(* IEC 61131-3 sources: guidance-for-physical-ai-production-designer-on-aws/source/plan2cell/crates/plan2cell/tests/fixtures/deploy_check/scene_fit/plc/codesys/head/GVL, 1 file *)

(* ---- GVL_Cell.st ---- *)
(*
 * GVL_Cell - generated by bt2plc 0.1.0 - DO NOT EDIT
 * Plan   : bt_1792156523_scene_fit (cell scene_fit)
 * Grants : planned ticket order
 * IL01   : R1#1 W02 > R2#2 W03 > R1#3 HOME
 * IL02   : R2#1 W01 > R1#2 W04 > R2#3 HOME
 *)
{attribute 'qualified_only'}
VAR_GLOBAL CONSTANT
    (* ========================================================================
       DIMENSIONS (array bounds are literals; *_DIM >= 1)
       ======================================================================== *)
    N_ROBOTS                : INT := 2;
    N_ZONES                 : INT := 2;
    N_OPS                   : INT := 6;
    N_PREDS                 : INT := 0;

    (* ========================================================================
       PROTOCOL / TIMING
       ======================================================================== *)
    PLAN_ID                 : WORD := WORD#16#A1BE;             (* fold of the plan fingerprint *)
    PROD_FOLGE              : WORD := WORD#11;                  (* default production Folge *)
    HOME_FOLGE              : WORD := WORD#125;                 (* blind homing *)
    JOB_NUMBER_BYTE         : BOOL := TRUE;                     (* FALSE: WORD LE bytes 2-3, TRUE: byte 2 *)
    PROFILE_VW              : BOOL := TRUE;                     (* TRUE: VW KS24 signal map and Folge handshake instead of the simulator telegram *)
    GRANT_POLICY            : E_GrantPolicy := E_GrantPolicy.GP_PLANNED;
    HOME_SEQUENTIAL         : BOOL := TRUE;
    AUTO_RUN                : BOOL := TRUE;                     (* start the next cycle automatically *)
    STEP_BYTE               : INT := 4;                         (* robot -> PLC, WORD LE op index *)
    REQ_BYTE                : INT := 28;                        (* robot -> PLC, DWORD LE zone requests *)
    GRANT_BYTE              : INT := 12;                        (* PLC -> robot, DWORD LE zone grants *)
    PLAN_ID_BYTE            : INT := 0;                         (* PLC -> robot, WORD LE plan id *)
    PERMIT_MASK             : DWORD := DWORD#16#80000000;       (* bit 31: permit predecessors *)
    T_RESET_PULSE           : TIME := T#1S;
    T_START_PULSE           : TIME := T#500MS;
    T_STOP_PULSE            : TIME := T#1S;
    T_HANDSHAKE             : TIME := T#5S;
    T_BRINGUP_LIMIT         : TIME := T#1M;                     (* safety enable: PROFINET connection set-up *)
    T_MISMATCH_DEBOUNCE     : TIME := T#200MS;
    T_STOP_DEBOUNCE         : TIME := T#200MS;                  (* job running: ProgRunning and ProgFinished low this long = robot stopped *)
    T_CYCLE_PAUSE           : TIME := T#2S;
    T_START_LIMIT           : TIME := T#15S;
    T_ABORT_LIMIT           : TIME := T#10S;
    T_HOME_LIMIT            : TIME := T#15S500MS;

    (* ========================================================================
       VW KS24 SIGNAL INDICES (used when PROFILE_VW; $IN/$OUT index, 1-based)
       ======================================================================== *)
    VW_READY_OUT            : INT := 9;                         (* O_R_Bereit *)
    VW_RK100_OUT            : INT := 10;                        (* O_R_RK100 safety circuit *)
    VW_AUTO_OUT             : INT := 12;                        (* O_R_Auto *)
    VW_ESTOP_OUT            : INT := 13;                        (* O_R_Notaus *)
    VW_END_OUT              : INT := 14;                        (* O_R_F_ENDE / LPKT *)
    VW_PF0_OUT              : INT := 15;                        (* O_R_PFO home position *)
    VW_STEP_OUT             : INT := 97;                        (* P_PktNr_SPS op index (16 bits) *)
    VW_REL_OUT              : INT := 41;                        (* interlock releases A41-56 *)
    VW_REQ_OUT              : INT := 81;                        (* interlock requests A81-96 *)
    VW_ERR_OUT              : INT := 225;                       (* VW_FEH_BIN_A error code (8 bits) *)
    VW_DRIVES_IN            : INT := 10;                        (* I_R_Ant_Ein *)
    VW_SRB_IN               : INT := 9;                         (* I_R_SRB Folge start *)
    VW_RESET_IN             : INT := 26;                        (* I_R_Quit_St acknowledge *)
    anInterlock             : ARRAY[1..4] OF INT := [1,2,1,2];  (* robot r, zone z -> VW interlock 1..16 (0 = not a member): index (r-1)*2+z *)

    (* ========================================================================
       ROBOTS (index = BT order)
       ======================================================================== *)
    asRobotTag              : ARRAY[1..2] OF STRING(16) := ['R1', 'R2'];
    asRobotNs               : ARRAY[1..2] OF STRING(32) := ['robot1', 'robot2'];
    abRobotActive           : ARRAY[1..2] OF BOOL := [TRUE, TRUE];
    abSafetyBypass          : ARRAY[1..2] OF BOOL := [FALSE, FALSE];(* SIMULATION ONLY: PROFIsafe slot-1 bits not required ([[robot]] safety_bypass) *)
    awRobotProdFolge        : ARRAY[1..2] OF WORD := [WORD#11, WORD#11];
    anRobotFirstOp          : ARRAY[1..2] OF INT := [1, 4];     (* op k of robot r: aOps[anRobotFirstOp[r] + k - 1] *)
    anRobotOpCount          : ARRAY[1..2] OF INT := [3, 3];

    (* ========================================================================
       ZONES - tickets of zone z: aTickets[anZoneFirst[z] .. anZoneFirst[z] + anZoneCount[z] - 1]
       ======================================================================== *)
    asZoneName              : ARRAY[1..2] OF STRING(8) := ['IL01', 'IL02'];
    anZoneFirst             : ARRAY[1..2] OF INT := [1, 4];
    anZoneCount             : ARRAY[1..2] OF INT := [3, 3];
    aTickets                : ARRAY[1..6] OF ST_Ticket := [
        (nRobot := 1, nOp := 1),    (* IL01 R1 #1 W02 *)
        (nRobot := 2, nOp := 2),    (* R2 #2 W03 *)
        (nRobot := 1, nOp := 3),    (* R1 #3 HOME *)
        (nRobot := 2, nOp := 1),    (* IL02 R2 #1 W01 *)
        (nRobot := 1, nOp := 2),    (* R1 #2 W04 *)
        (nRobot := 2, nOp := 3)    (* R2 #3 HOME *)
    ];

    (* ========================================================================
       OPS - op k of robot r: aOps[anRobotFirstOp[r] + k - 1]
       ======================================================================== *)
    (* tLimit = 1.5 x tExpected + 5 s ; tZoneDeadline = 1.5 x ASAP grant + (5 + 0.2) s x depth + 10 s *)
    aOps                    : ARRAY[1..6] OF ST_OpInfo := [
        (nRobot := 1, nOp := 1, dwZoneMask := DWORD#16#00000001, nPredFirst := 0, nPredCount := 0, tExpected := T#7S408MS, tLimit := T#16S112MS, tZoneDeadline := T#10S, sName := 'W02'),    (* R1 #1 W02 *)
        (nRobot := 1, nOp := 2, dwZoneMask := DWORD#16#00000002, nPredFirst := 0, nPredCount := 0, tExpected := T#5S118MS, tLimit := T#12S677MS, tZoneDeadline := T#33S680MS, sName := 'W04'),    (* R1 #2 W04 *)
        (nRobot := 1, nOp := 3, dwZoneMask := DWORD#16#00000001, nPredFirst := 0, nPredCount := 0, tExpected := T#4S522MS, tLimit := T#11S783MS, tZoneDeadline := T#46S557MS, sName := 'HOME'),    (* R1 #3 HOME *)
        (nRobot := 2, nOp := 1, dwZoneMask := DWORD#16#00000002, nPredFirst := 0, nPredCount := 0, tExpected := T#12S320MS, tLimit := T#23S480MS, tZoneDeadline := T#10S, sName := 'W01'),    (* R2 #1 W01 *)
        (nRobot := 2, nOp := 2, dwZoneMask := DWORD#16#00000001, nPredFirst := 0, nPredCount := 0, tExpected := T#5S117MS, tLimit := T#12S676MS, tZoneDeadline := T#33S680MS, sName := 'W03'),    (* R2 #2 W03 *)
        (nRobot := 2, nOp := 3, dwZoneMask := DWORD#16#00000002, nPredFirst := 0, nPredCount := 0, tExpected := T#10S293MS, tLimit := T#20S440MS, tZoneDeadline := T#46S557MS, sName := 'HOME')    (* R2 #3 HOME *)
    ];

    (* ========================================================================
       PERMIT PREDECESSORS - op preds: aPreds[nPredFirst .. nPredFirst + nPredCount - 1]
       ======================================================================== *)
    aPreds                  : ARRAY[1..1] OF ST_Ticket := [
        (nRobot := 0, nOp := 0)    (* no permit predecessors *)
    ];
END_VAR
